TYPE T_ServiceTimeHandle : UDINT;
END_TYPE

(* stored: Version 1.1.0.1, ProductVersion 3.1.4026.18
   DUT T_ServiceTimeHandle: Id {3b37d66e-5422-437a-b01b-eae2c52fd5a4} *)
